# EPICS substitutions: iocs/motor/aerotech-ioc/db/Ensemble.substitutions
# C's iocAerotech Ensemble.substitutions, P and PORT from st.cmd.
file "$(MOTOR)/db/asyn_motor.db"
{
pattern
{N,  M,       DTYP,         ADDR,  DESC,          EGU,  DIR,  VELO,  VBAS,  ACCL,  BDST,  BVEL,  BACC,  MRES,     PREC,  DHLM,  DLLM,  INIT}
{1,  "m$(N)", "asynMotor",  0,     "motor $(N)",  mm,   Pos,  .1,    0,     .2,    0,     1,     .2,    1.25E-5,  7,     0,     0,     "SCURVE 100"}
}
